Fanuc KAREL source: KA00197.KL

PROGRAM KA00197
%NOLOCKGROUP
VAR
  SRC: ARRAY[4] OF SHORT
  DST: ARRAY[4] OF XYZWPR
BEGIN
  DST = SRC
END KA00197
